FUNCTION_BLOCK DestinationTypeMismatch
  (* Standard: 61499-1; Description: Copyright (c) 2026 Martin Erich Jobst This program and the accompanying materials are made available under the terms of the Eclipse Public License 2.0 which is available at https://www.eclipse.org/legal/epl-2.0/ SPDX-License-Identifier: EPL-2.0 *)
  (* Version 1.0, 2026-11-18, Martin Jobst *)
  PACKAGE lib::VarDeclaration;
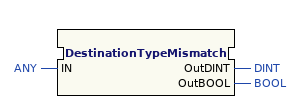
  VAR_INPUT
    IN : ANY;
  END_VAR
  VAR_OUTPUT
    OutDINT : DINT;
    OutBOOL : BOOL;
  END_VAR
  DATA_CONNECTIONS
    IN TO OutDINT;
    IN TO OutBOOL;
  END_CONNECTIONS
END_FUNCTION_BLOCK
